// TIA Portal V19 export
VAR_GLOBAL   // PLC tag table "Spare"
   "DI_Spare_I1.3" AT %I1.3 : Bool;
   "DI_Spare_I1.4" AT %I1.4 : Bool;
   "DI_Spare_I1.5" AT %I1.5 : Bool;
   "DQ_Spare_Q1.0" AT %Q1.0 : Bool;
   "DQ_Spare_Q1.1" AT %Q1.1 : Bool;
   "DI_Spare_I8.5" AT %I8.5 : Bool;
   "DI_Spare_I8.6" AT %I8.6 : Bool;
   "DI_Spare_I8.7" AT %I8.7 : Bool;
   "DI_Spare_I9.0" AT %I9.0 : Bool;
   "DI_Spare_I9.1" AT %I9.1 : Bool;
   "DI_Spare_I9.2" AT %I9.2 : Bool;
   "DI_Spare_I9.3" AT %I9.3 : Bool;
   "DI_Spare_I9.4" AT %I9.4 : Bool;
   "DI_Spare_I9.5" AT %I9.5 : Bool;
   "DI_Spare_I9.6" AT %I9.6 : Bool;
   "DI_Spare_I9.7" AT %I9.7 : Bool;
   "DI_Spare_I13.7" AT %I13.7 : Bool;
   "DQ_Spare_Q17.7" AT %Q17.7 : Bool;
   "DI_Spare_I1.2" AT %I1.2 : Bool;
END_VAR
